(* PLC project PR_FibroMainSeq_Soft2.0 1_workflow_a30ae2_PLC, SiemensToBackhoff Siemens TIA Portal → Beckhoff TwinCAT PLCopen Converter 2.2 *)
(* stored: creationDateTime 2026-10-12T12:22:45.841201, modificationDateTime 2026-10-12T12:22:45.841201 *)

FUNCTION_BLOCK PR_FibroMainSeq_Soft2.0 1_workflow_a30ae2
VAR_INPUT
	iAllStationsSafe : BOOL;
	iAllTaskOver : BOOL;
	iAutoRunning : BOOL;
	iFaultReset : BOOL;
	iFibroAtStnPos : BOOL;
	iIndexOver : BOOL;
	iProcessActive : BOOL;
	iReset_fault : BOOL;
	iSstMode : BOOL;
	iSstPB : BOOL;
END_VAR
VAR_OUTPUT
	qError : ARRAY[1..1] OF BOOL;
	qMessage_0 : BOOL;
	qProcessActive : BOOL;
END_VAR
VAR
	c10_ChkRecCond_T1 : BOOL;
	c10_ChkRecCond_T2 : BOOL;
	c10_ChkRecCond_T3 : BOOL;
	c50_ChkPartPresentAtStn_T1 : BOOL;
	c50_ChkPartPresentAtStn_T2 : BOOL;
	StateNo : INT;
	s100_WtAllStnTaskOver : BOOL;
	s100_WtAllStnTaskOver_T1 : BOOL;
	s10_ChkRecCond : BOOL;
	s10_ChkRecCond_T1 : BOOL;
	s10_ChkRecCond_T2 : BOOL;
	s10_ChkRecCond_T3 : BOOL;
	s130_ChkAllStnSafe2 : BOOL;
	s130_ChkAllStnSafe2_T1 : BOOL;
	s140_WtIndexOver : BOOL;
	s140_WtIndexOver_T1 : BOOL;
	s1_WtResetRel : BOOL;
	s1_WtResetRel_T1 : BOOL;
	s20_WtManualIntv : BOOL;
	s20_WtManualIntv_T1 : BOOL;
	s30_WtFibroAtStnPos : BOOL;
	s30_WtFibroAtStnPos_T1 : BOOL;
	s40_ChkAllStnSafe : BOOL;
	s40_ChkAllStnSafe_T1 : BOOL;
	s50_ChkPartPresentAtStn : BOOL;
	s50_ChkPartPresentAtStn_T1 : BOOL;
	s50_ChkPartPresentAtStn_T2 : BOOL;
	s60_WtPartPresentAtStn : BOOL;
	s60_WtPartPresentAtStn_T1 : BOOL;
	sAbnormalCondition : BOOL;
	sPartPresentAtStation : BOOL;
	sProcessActive : BOOL;
	sSst : BOOL;
	sSstPulse : BOOL;
	sSstRise : R_TRIG;
	sStWtResetRel : BOOL;
	sStWtResetRel_T1 : BOOL;
END_VAR
VAR_TEMP
	tOne : BOOL;
END_VAR
  VAR  (* added by the conversion: wires and edge detectors of the diagram *)
    _w24 : BOOL;
    _w26 : BOOL;
    _w39 : BOOL;
    _w41 : BOOL;
    _w42 : BOOL;
    _w74 : BOOL;
    _w78 : BOOL;
    _w79 : BOOL;
    _w80 : BOOL;
    _w81 : BOOL;
    _w94 : BOOL;
    _w96 : BOOL;
    _w97 : BOOL;
    _w114 : BOOL;
    _w116 : BOOL;
    _w117 : BOOL;
    _w135 : BOOL;
    _w137 : BOOL;
    _w138 : BOOL;
    _w162 : BOOL;
    _w164 : BOOL;
    _w165 : BOOL;
    _w166 : BOOL;
    _w180 : BOOL;
    _w182 : BOOL;
    _w183 : BOOL;
    _w196 : BOOL;
    _w200 : BOOL;
    _w201 : BOOL;
    _w218 : BOOL;
    _w220 : BOOL;
    _w221 : BOOL;
    _w238 : BOOL;
    _w240 : BOOL;
    _w241 : BOOL;
  END_VAR

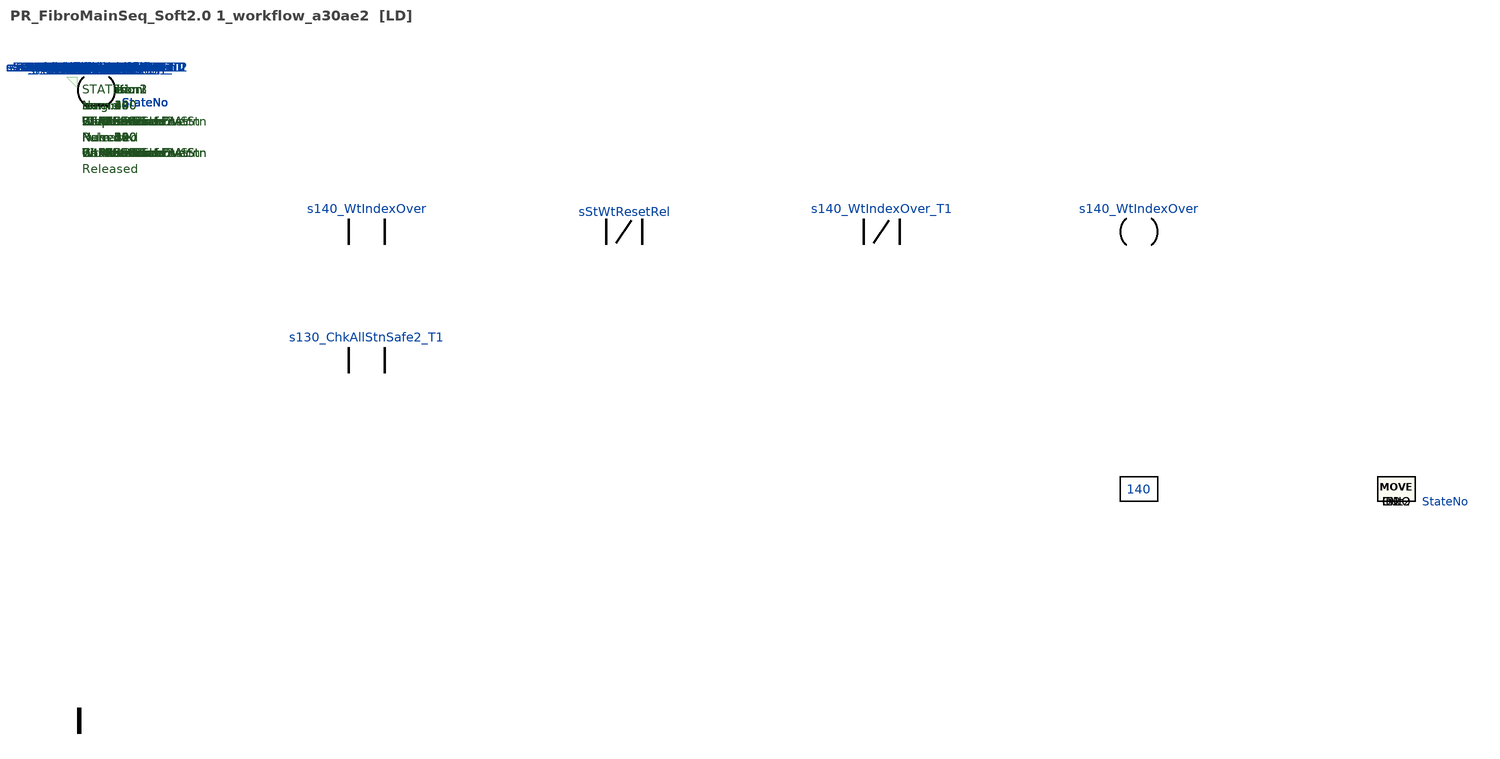
(* LD diagram, written out as Structured Text *)
(* Network 1 *)
(* Create Single Step Pulse bit *)
(* Create Single Step bit *)
(* Transition for STATE Num:0 Reset Released *)
(* STATE Num:0 Reset Released *)
(* Transition for STATE Num:1 WtResetRel *)
(* STATE Num:1 WtResetRel *)
(* Condition1 for STATE Num:10 ChkRecCond *)
(* Condition2 for STATE Num:10 ChkRecCond *)
(* Condition3 for STATE Num:10 ChkRecCond *)
(* Transition for STATE Num:10 ChkRecCond *)
(* STATE Num:10 ChkRecCond *)
(* Transition for STATE Num:20 WtManualIntv *)
(* STATE Num:20 WtManualIntv *)
(* Actions for STATE Num:20 WtManualIntv *)
(* Transition for STATE Num:40 ChkAllStnSafe *)
(* STATE Num:40 ChkAllStnSafe *)
(* Actions for STATE Num:40 ChkAllStnSafe *)
(* Transition for STATE Num:30 WtFibroAtStnPos *)
(* STATE Num:30 WtFibroAtStnPos *)
(* Condition1 for STATE Num:50 ChkPartPresentAtStn *)
(* Condition2 for STATE Num:50 ChkPartPresentAtStn *)
(* Transition for STATE Num:50 ChkPartPresentAtStn *)
(* STATE Num:50 ChkPartPresentAtStn *)
(* Transition for STATE Num:60 WtPartPresentAtStn *)
(* STATE Num:60 WtPartPresentAtStn *)
(* Transition for STATE Num:100 WtAllStnTaskOver *)
(* STATE Num:100 WtAllStnTaskOver *)
(* Actions for STATE Num:100 WtAllStnTaskOver *)
(* Transition for STATE Num:130 ChkAllStnSafe2 *)
(* STATE Num:130 ChkAllStnSafe2 *)
(* Actions for STATE Num:130 ChkAllStnSafe2 *)
(* Transition for STATE Num:140 WtIndexOver *)
(* STATE Num:140 WtIndexOver *)
tOne := tOne OR NOT tOne;
sSstRise(CLK := iSstPB);
sSstPulse := sSstRise.Q;
sSst := iSstMode AND sSstPulse OR NOT iSstMode;
sStWtResetRel_T1 := sStWtResetRel AND iAutoRunning;
_w24 := sStWtResetRel;
_w26 := (_w24 OR NOT iAutoRunning) AND NOT sStWtResetRel_T1;
sStWtResetRel := _w26;
IF _w26 THEN StateNo := 0; END_IF;
s1_WtResetRel_T1 := s1_WtResetRel AND NOT sStWtResetRel AND sSst AND iAutoRunning;
_w39 := s1_WtResetRel;
_w41 := (_w39 OR sStWtResetRel_T1) AND NOT sStWtResetRel;
_w42 := _w41 AND NOT s1_WtResetRel_T1;
s1_WtResetRel := _w42;
IF _w42 THEN StateNo := 1; END_IF;
c10_ChkRecCond_T1 := sAbnormalCondition;
c10_ChkRecCond_T2 := iProcessActive;
c10_ChkRecCond_T3 := NOT iProcessActive;
s10_ChkRecCond_T1 := s10_ChkRecCond AND NOT sStWtResetRel AND sSst AND c10_ChkRecCond_T1;
s10_ChkRecCond_T2 := s10_ChkRecCond AND NOT sStWtResetRel AND sSst AND NOT s10_ChkRecCond_T1 AND c10_ChkRecCond_T2;
s10_ChkRecCond_T3 := s10_ChkRecCond AND NOT sStWtResetRel AND sSst AND NOT s10_ChkRecCond_T1 AND NOT s10_ChkRecCond_T1 AND NOT s10_ChkRecCond_T2 AND c10_ChkRecCond_T3;
_w74 := s10_ChkRecCond;
_w78 := (_w74 OR s1_WtResetRel_T1 OR s20_WtManualIntv_T1 OR s140_WtIndexOver_T1) AND NOT sStWtResetRel;
_w79 := _w78 AND NOT s10_ChkRecCond_T1;
_w80 := _w79 AND NOT s10_ChkRecCond_T2;
_w81 := _w80 AND NOT s10_ChkRecCond_T3;
s10_ChkRecCond := _w81;
IF _w81 THEN StateNo := 10; END_IF;
s20_WtManualIntv_T1 := s20_WtManualIntv AND NOT sStWtResetRel AND sSst AND iFaultReset;
_w94 := s20_WtManualIntv;
_w96 := (_w94 OR s10_ChkRecCond_T1) AND NOT sStWtResetRel;
_w97 := _w96 AND NOT s20_WtManualIntv_T1;
s20_WtManualIntv := _w97;
IF _w97 THEN StateNo := 20; END_IF;
qError[1] := s20_WtManualIntv;
s40_ChkAllStnSafe_T1 := s40_ChkAllStnSafe AND NOT sStWtResetRel AND sSst AND iAllStationsSafe;
_w114 := s40_ChkAllStnSafe;
_w116 := (_w114 OR s10_ChkRecCond_T3) AND NOT sStWtResetRel;
_w117 := _w116 AND NOT s40_ChkAllStnSafe_T1;
s40_ChkAllStnSafe := _w117;
IF _w117 THEN StateNo := 40; END_IF;
qMessage_0 := s40_ChkAllStnSafe;
s30_WtFibroAtStnPos_T1 := s30_WtFibroAtStnPos AND NOT sStWtResetRel AND sSst AND (iFibroAtStnPos OR iIndexOver);
_w135 := s30_WtFibroAtStnPos;
_w137 := (_w135 OR s40_ChkAllStnSafe_T1) AND NOT sStWtResetRel;
_w138 := _w137 AND NOT s30_WtFibroAtStnPos_T1;
s30_WtFibroAtStnPos := _w138;
IF _w138 THEN StateNo := 30; END_IF;
c50_ChkPartPresentAtStn_T1 := NOT sPartPresentAtStation;
c50_ChkPartPresentAtStn_T2 := sPartPresentAtStation;
s50_ChkPartPresentAtStn_T1 := s50_ChkPartPresentAtStn AND NOT sStWtResetRel AND sSst AND c50_ChkPartPresentAtStn_T1;
s50_ChkPartPresentAtStn_T2 := s50_ChkPartPresentAtStn AND NOT sStWtResetRel AND sSst AND NOT s50_ChkPartPresentAtStn_T1 AND c50_ChkPartPresentAtStn_T2;
_w162 := s50_ChkPartPresentAtStn;
_w164 := (_w162 OR s30_WtFibroAtStnPos_T1) AND NOT sStWtResetRel;
_w165 := _w164 AND NOT s50_ChkPartPresentAtStn_T1;
_w166 := _w165 AND NOT s50_ChkPartPresentAtStn_T2;
s50_ChkPartPresentAtStn := _w166;
IF _w166 THEN StateNo := 50; END_IF;
s60_WtPartPresentAtStn_T1 := s60_WtPartPresentAtStn AND NOT sStWtResetRel AND sSst AND sPartPresentAtStation AND iAllStationsSafe;
_w180 := s60_WtPartPresentAtStn;
_w182 := (_w180 OR s50_ChkPartPresentAtStn_T1) AND NOT sStWtResetRel;
_w183 := _w182 AND NOT s60_WtPartPresentAtStn_T1;
s60_WtPartPresentAtStn := _w183;
IF _w183 THEN StateNo := 60; END_IF;
s100_WtAllStnTaskOver_T1 := s100_WtAllStnTaskOver AND NOT sStWtResetRel AND sSst AND iAllTaskOver;
_w196 := s100_WtAllStnTaskOver;
_w200 := (_w196 OR s10_ChkRecCond_T2 OR s50_ChkPartPresentAtStn_T2 OR s60_WtPartPresentAtStn_T1) AND NOT sStWtResetRel;
_w201 := _w200 AND NOT s100_WtAllStnTaskOver_T1;
s100_WtAllStnTaskOver := _w201;
IF _w201 THEN StateNo := 100; END_IF;
qProcessActive := s100_WtAllStnTaskOver;
s130_ChkAllStnSafe2_T1 := s130_ChkAllStnSafe2 AND NOT sStWtResetRel AND sSst AND iAllStationsSafe;
_w218 := s130_ChkAllStnSafe2;
_w220 := (_w218 OR s100_WtAllStnTaskOver_T1) AND NOT sStWtResetRel;
_w221 := _w220 AND NOT s130_ChkAllStnSafe2_T1;
s130_ChkAllStnSafe2 := _w221;
IF _w221 THEN StateNo := 130; END_IF;
qMessage_0 := s130_ChkAllStnSafe2;
s140_WtIndexOver_T1 := s140_WtIndexOver AND NOT sStWtResetRel AND sSst AND iIndexOver;
_w238 := s140_WtIndexOver;
_w240 := (_w238 OR s130_ChkAllStnSafe2_T1) AND NOT sStWtResetRel;
_w241 := _w240 AND NOT s140_WtIndexOver_T1;
s140_WtIndexOver := _w241;
IF _w241 THEN StateNo := 140; END_IF;
END_FUNCTION_BLOCK
